DATA_BLOCK "GDB_IoBridgeEpoch"
{ S7_Optimized_Access := 'TRUE' }
VERSION : 0.1
RETAIN
VAR
    Epoch {ExternalAccessible := 'False'; ExternalVisible := 'False'; ExternalWritable := 'False'} : UDInt;
END_VAR
BEGIN
END_DATA_BLOCK
